TYPE "FRK_Profiler_DeclarationUnit"
VERSION : 0.1
   STRUCT
      LastCycle : "FRK_CycleProfile_DeclarationUnit";
      StepStats : Array[1..4] of "ST_TimingRow";
      StatsTruncated : Bool;
      LastCycleTime : Time;
      MinCycleTime : Time;
      History : Array[1..60] of "ST_CycleSummary";
      HistoryHead : Int;
   END_STRUCT;

END_TYPE

